Fanuc KAREL source: kt00611.KL

-- PROVISIONAL review KL for V1013-1; original PC SHA256 e1eb27336adcb42f18bbe4a895694992c060f875e2c151aa1fc286656520a327
-- Incomplete behavior may be omitted. Consult companion uncertainty JSON. Do not deploy.
PROGRAM KT00611
%NOLOCKGROUP
VAR
  R1 : REAL
  R2 : REAL
  OUT : REAL
BEGIN
  -- UNRESOLVED_PC offsets 5-16; opcodes 2E,23
  -- UNRESOLVED_PC offsets 21-32; opcodes 2E,23
  -- UNRESOLVED_PC offsets 37-48; opcodes 2E,23
  -- UNRESOLVED_PC offsets 53-64; opcodes 2E,23
  -- UNRESOLVED_PC offsets 69-81; opcodes 21,23
  -- UNRESOLVED_PC offsets 86-90; opcodes 7F
END KT00611
